// TIA Portal V20 export
// export: Created 2026-10-12T05:42:33.5214407Z, ExportSetting WithDefaults, DisplayName Totally Integrated Automation Portal, DisplayVersion V20, DisplayName TIA Portal Openness, DisplayVersion V20, DisplayName TIA Portal Teamcenter Gateway, DisplayVersion V20, DisplayName TIA Portal Version Control Interface, DisplayVersion V20, DisplayName SINAMICS Startdrive Advanced, DisplayVersion V20 SP1 Update 2, DisplayName SINAMICS Startdrive G110M, G120, G120C, G120D, G120P, G115D, DisplayVersion V20 SP1 Update 2, DisplayName SINAMICS Startdrive G130, G150, S120, S150, SINAMICS MV, G220, S200, S210, DisplayVersion V20 SP1 Update 2, DisplayName STEP 7 Professional, DisplayVersion V20, DisplayName STEP 7 Safety, DisplayVersion V20, DisplayName WinCC Basic/Comfort/Advanced, DisplayVersion V20, DisplayName WinCC Professional, DisplayVersion V20, DisplayName WinCC Unified, DisplayVersion V20
FUNCTION "F_CylinderSequenceLease" : Void   // FC156, SCL
{ S7_Optimized_Access := 'TRUE' }
VERSION : 0.1
// stored: AutoNumber true, IsIECCheckEnabled false, SetENOAutomatically false, UDAEnableTagReadback false
   VAR_IN_OUT
      Seq : "FRK_SequenceCtx";
      Target : "FB_CylinderCM";
   END_VAR
BEGIN

   IF #Target.Device.Lease.OwnerIndex = #Seq.OwnerIndex
       AND #Target.Device.Lease.ChainIndex = #Seq.ChainIndex
       AND #Target.Device.Lease.BranchIndex = #Seq.BranchIndex
       AND #Seq.OwnerIndex > 0 AND #Seq.ChainIndex > 0
       AND (NOT #Seq.Running OR #Seq.Error OR #Seq.Restart) THEN
       #Target.Device.Withdrawn := TRUE;
   END_IF;
   IF #Target.Device.Lease.OwnerIndex = #Seq.OwnerIndex
       AND #Target.Device.Lease.ChainIndex = #Seq.ChainIndex
       AND #Target.Device.Lease.BranchIndex = #Seq.BranchIndex
       AND #Target.Device.Lease.AbortIssued AND #Target.Device.Lease.ReleasedScan <> #Seq.Scan THEN
       #Target.Abort := FALSE;
       #Target.Device.Lease.AbortIssued := FALSE;
   END_IF;
   IF #Target.Device.Lease.Raised AND #Target.Device.Lease.OwnerIndex = #Seq.OwnerIndex
       AND #Target.Device.Lease.ChainIndex = #Seq.ChainIndex
       AND #Target.Device.Lease.BranchIndex = #Seq.BranchIndex
       AND (NOT #Seq.Running OR #Seq.Error OR #Seq.Restart OR #Target.Device.Lease.Step <> #Seq.Step) THEN
       #Target.Abort := #Target.Busy;
       #Target.Device.Lease.AbortIssued := #Target.Busy;
   END_IF;
   "FRK_SeqLease"(Seq := #Seq,
                  Lease := #Target.Device.Lease,
                  Execute := #Target.Execute);
END_FUNCTION
